(* IEC 61131-3 sources: avi-aoi-management/scripts/ai-eval/ngau-nhien/kho/st-tt5-crc16-modbus/khung/src, 1 file *)

(* ---- Crc16Modbus.st ---- *)
FUNCTION Crc16Modbus : WORD
VAR_INPUT
    DU_LIEU : ARRAY[0..63] OF BYTE;
    DO_DAI : INT;
END_VAR
    (* TODO: cài đặt theo đề bài *)
    Crc16Modbus := 0;
END_FUNCTION
